(*
SPDX-FileCopyrightText: © 2026 Oleksandr Tiutyk <trofimich@gmail.com>
SPDX-License-Identifier: MIT
License: https://opensource.org/license/mit
*)

(*!
<summary>Beckhoff EL5152 32-bit incremental encoder feedback without a latch.</summary>
<description>
Represents the 32-bit main input PDO for one EL5152 channel (0x1A00 or 0x1A04).
Status is 16-bit; Value is the 32-bit counter. This terminal has no latch value.
Optional period/frequency PDOs are outside this channel; disable them or link them separately.
Link fields individually and evaluate bus/channel validity before use; unlinked zeros are not valid data.
Use one owner task and externally synchronize other access. Copies are not atomic multi-field snapshots.
When used for I/O, link located fields or their containing buffers to the matching selected PDOs.
The record is not a packed wire buffer; compiler padding is not part of the device specification.
Unlinked/default values do not prove valid I/O. The caller evaluates bus/channel validity before use.
Use one owner task per instance and externally synchronize other access; multi-field snapshots are not atomic.
Copies store data without creating hardware links. Keep borrowed field references valid while consumers are bound.
This passive record performs no validation, synchronization, configuration or protocol advancement.
</description>
*)
TYPE INCREMENTAL_ENCODER_COUNTER_INPUT_CHANNEL :
STRUCT
	Status AT %I* : WORD;
	Value AT %I* : UDINT;
END_STRUCT
END_TYPE

(* stored: Version 1.1.0.1
   DUT INCREMENTAL_ENCODER_COUNTER_INPUT_CHANNEL: Id {29f09c50-d0c9-46aa-9f0c-045dd35af63c} *)
